Fanuc KAREL source: KT00548.KL

PROGRAM KT00548
%NOLOCKGROUP
VAR
  P1: JOINTPOS
  P2: JOINTPOS
  OUT: BOOLEAN
BEGIN
  OUT = P1 >=< P2
END KT00548
